Fanuc KAREL source: KA00026.KL

PROGRAM KA00026
%NOLOCKGROUP
VAR
  SRC: BOOLEAN
  DST: REAL
BEGIN
  SRC = TRUE
  DST = SRC
END KA00026
